FUNCTION_BLOCK supervision (* Extracted Composite Function Block Type *)
  (* Standard: 61499-2 *)
  (* Version 10/27/2026, lizar *)
  PACKAGE Main;
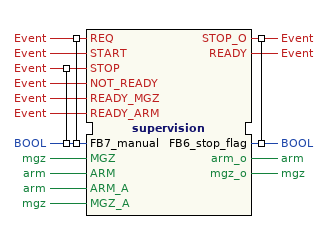
  EVENT_INPUT
    REQ WITH FB7_manual; (* Initialization Request *)
    START; (* Initialization Request *)
    STOP WITH FB7_manual;
    NOT_READY; (* Reset Event *)
    READY_MGZ; (* Second Event Input *)
    READY_ARM; (* First Event Input *)
  END_EVENT
  EVENT_OUTPUT
    STOP_O WITH FB6_stop_flag; (* Execution Confirmation *)
    READY; (* Rendezvous Output Event *)
  END_EVENT
  VAR_INPUT
    FB7_manual : BOOL;
  END_VAR
  VAR_OUTPUT
    FB6_stop_flag : BOOL; (* Output event qualifier *)
  END_VAR
  SOCKETS
    MGZ : mgz;
    ARM : arm;
    ARM_A : arm;
    MGZ_A : mgz;
  END_SOCKETS
  PLUGS
    arm_o : arm;
    mgz_o : mgz;
  END_PLUGS
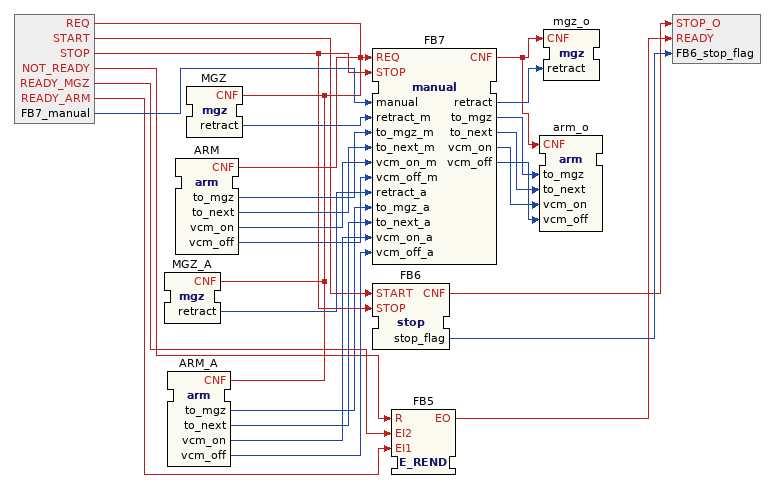
  FBS
    FB5 : E_REND;
    FB6 : stop;
    FB7 : manual;
  END_FBS
  EVENT_CONNECTIONS
    START TO FB6.START;
    FB6.CNF TO STOP_O;
    REQ TO FB7.REQ;
    STOP TO FB7.STOP;
    NOT_READY TO FB5.R;
    READY_MGZ TO FB5.EI2;
    READY_ARM TO FB5.EI1;
    FB5.EO TO READY;
    STOP TO FB6.STOP;
    MGZ.CNF TO FB7.REQ;
    ARM.CNF TO FB7.REQ;
    ARM_A.CNF TO FB7.REQ;
    MGZ_A.CNF TO FB7.REQ;
    FB7.CNF TO arm_o.CNF;
    FB7.CNF TO mgz_o.CNF;
  END_CONNECTIONS
  DATA_CONNECTIONS
    FB6.stop_flag TO FB6_stop_flag;
    FB7_manual TO FB7.manual;
    MGZ.retract TO FB7.retract_m;
    ARM.to_mgz TO FB7.to_mgz_m;
    ARM.to_next TO FB7.to_next_m;
    ARM.vcm_on TO FB7.vcm_on_m;
    ARM.vcm_off TO FB7.vcm_off_m;
    ARM_A.to_mgz TO FB7.to_mgz_a;
    ARM_A.to_next TO FB7.to_next_a;
    ARM_A.vcm_on TO FB7.vcm_on_a;
    ARM_A.vcm_off TO FB7.vcm_off_a;
    MGZ_A.retract TO FB7.retract_a;
    FB7.to_mgz TO arm_o.to_mgz;
    FB7.to_next TO arm_o.to_next;
    FB7.vcm_on TO arm_o.vcm_on;
    FB7.vcm_off TO arm_o.vcm_off;
    FB7.retract TO mgz_o.retract;
  END_CONNECTIONS
END_FUNCTION_BLOCK
